Fanuc KAREL source: kb00146.compact.KL

PROGRAM KB00146
%STACKSIZE=65535
%PRIORITY=65535
%NOLOCKGROUP
%ENVIRONMENT FDEV
VAR
P1 : STRING[80]
P2 : STRING[80]
P3 : BOOLEAN
P4 : INTEGER
BEGIN
P1='A'
P2='A'
P3=TRUE
P4=1
RENAME_FILE(P1,P2,P3,P4)
END KB00146
